DATA_BLOCK "naut_SfcAssocForms_DB"
{ S7_Optimized_Access := 'TRUE' }
VERSION : 0.1
"naut_SfcAssocForms"

BEGIN

END_DATA_BLOCK
